// TIA Portal project "IncrocioSemaforicoT" (V19)

(* hardware
DEVICE "S7-1200 station_1"  S7-1200 Station
   slot 0: "Rack_0"  S7-1200 Rack  Rack  V1.0
   slot 1: "PLC_1"  CPU 1212C DC/DC/Rly  6ES7 212-1HE40-0XB0  V4.6
   slot 2: "DQ 16x24VDC_1"  SM 1222 DQ16 x 24VDC  6ES7 222-1BH32-0XB0  V2.0
DEVICE "HMI_1"  KTP700 Basic PN
   slot 0: "HMI_1"  KTP700 Basic PN  6AV2 123-2GB03-0AX0  17.0.0.0
   slot 1: "HMI_RT_1"  KTP700 Basic PN  6AV2 123-2GB03-0AX0  17.0.0.0
   slot 5: "HMI_1.IE_CP_1"  PROFINET Interface  17.0.0.0
      slot 1: "PROFINET Interface_1"  PROFINET Interface
         slot 1: "Port_1"  Port
*)

// ===== PLC "PLC_1"  CPU 1212C DC/DC/Rly =====

VAR_GLOBAL   // PLC tag table "Default tag table"
   "PulsantePedonale1" AT %I0.0 : Bool;
   "PulsantePedonale2" AT %I0.1 : Bool;
   "PulsantePedonale3" AT %I0.2 : Bool;
   "VerdePedonale1" AT %Q0.3 : Bool;
   "GialloPedonale1" AT %Q0.6 : Bool;
   "RossoVeicolare1" AT %Q1.1 : Bool;
   "VerdeVeicolare1" AT %Q1.4 : Bool;
   "GialloVeicolare1" AT %Q1.7 : Bool;
   "RossoPedonale1" AT %Q0.0 : Bool;
   "RossoPedonale2" AT %Q0.1 : Bool;
   "RossoPedonale3" AT %Q0.2 : Bool;
   "VerdePedonale2" AT %Q0.4 : Bool;
   "VerdePedonale3" AT %Q0.5 : Bool;
   "GialloPedonale2" AT %Q0.7 : Bool;
   "GialloPedonale3" AT %Q1.0 : Bool;
   "RossoVeicolare2" AT %Q1.2 : Bool;
   "RossoVeicolare3" AT %Q1.3 : Bool;
   "VerdeVeicolare2" AT %Q1.5 : Bool;
   "VerdeVeicolare3" AT %Q1.6 : Bool;
   "GialloVeicolare2" AT %Q2.0 : Bool;
   "GialloVeicolare3" AT %Q2.1 : Bool;
   "AppoggioGialloVeicolare1" AT %M0.0 : Bool;
   "AppoggioVerdeVeicolare1" AT %M0.1 : Bool;
   "AppoggioQTPRossoVeicolare1" AT %M0.2 : Bool;
   "AppoggioVerdeVeicolare2" AT %M0.3 : Bool;
   "AppoggioGialloVeicolare2" AT %M0.4 : Bool;
   "AppoggioQTPRossoVeicolare2" AT %M0.5 : Bool;
   "AppoggioVerdeVeicolare3" AT %M0.6 : Bool;
   "AppoggioGialloVeicolare3" AT %M0.7 : Bool;
   "AppoggioPulsante1" AT %M1.0 : Bool;
   "AppoggioPulsante2" AT %M1.1 : Bool;
   "AppoggioPulsante3" AT %M1.2 : Bool;
   "AppoggioNVerdePedonale1" AT %M1.3 : Bool;
   "RichiestaPedonale1" AT %M1.4 : Bool;
   "RichiestaPedonale2" AT %M1.5 : Bool;
   "RichiestaPedonale3" AT %M1.6 : Bool;
   "AppoggioPVerdePedonale1" AT %M1.7 : Bool;
   "AppoggioPVerdePedonale2" AT %M2.0 : Bool;
   "AppoggioPVerdePedonale3" AT %M2.1 : Bool;
   "AppoggioQTPRossoVeicolare3" AT %M2.2 : Bool;
   "AppoggioNVerdePedonale2" AT %M2.3 : Bool;
   "AppoggioNVerdePedonale3" AT %M2.4 : Bool;
   "AppoggioQTPRossoVeicolare1Pedonale1" AT %M2.5 : Bool;
   "AppoggioQTPRossoVeicolare1Pedonale3" AT %M2.6 : Bool;
   "AppoggioQTPRossoVeicolare2Pedonale1" AT %M2.7 : Bool;
   "AppoggioQTPRossoVeicolare2Pedonale2" AT %M3.0 : Bool;
   "AppoggioQTPRossoVeicolare3Pedonale2" AT %M3.1 : Bool;
   "AppoggioQTPRossoVeicolare3Pedonale3" AT %M3.2 : Bool;
END_VAR

// folder: System blocks/Program resources

DATA_BLOCK "TPRossoVeicolare1"   // DB1
{ S7_Optimized_Access := 'TRUE' }
AUTHOR : Simatic
FAMILY : IEC
NAME : IEC_TMR
VERSION : 1.0
// stored: InstanceOfName IEC_TIMER
"IEC_TIMER"
BEGIN
END_DATA_BLOCK

DATA_BLOCK "TPVerdeVeicolare1"   // DB2
{ S7_Optimized_Access := 'TRUE' }
AUTHOR : Simatic
FAMILY : IEC
NAME : IEC_TMR
VERSION : 1.0
// stored: InstanceOfName IEC_TIMER
"IEC_TIMER"
BEGIN
END_DATA_BLOCK

DATA_BLOCK "TPGialloVeicolare1"   // DB3
{ S7_Optimized_Access := 'TRUE' }
AUTHOR : Simatic
FAMILY : IEC
NAME : IEC_TMR
VERSION : 1.0
// stored: InstanceOfName IEC_TIMER
"IEC_TIMER"
BEGIN
END_DATA_BLOCK

DATA_BLOCK "TPVerdeVeicolare2"   // DB4
{ S7_Optimized_Access := 'TRUE' }
AUTHOR : Simatic
FAMILY : IEC
NAME : IEC_TMR
VERSION : 1.0
// stored: InstanceOfName IEC_TIMER
"IEC_TIMER"
BEGIN
END_DATA_BLOCK

DATA_BLOCK "TPGialloVeicolare2"   // DB5
{ S7_Optimized_Access := 'TRUE' }
AUTHOR : Simatic
FAMILY : IEC
NAME : IEC_TMR
VERSION : 1.0
// stored: InstanceOfName IEC_TIMER
"IEC_TIMER"
BEGIN
END_DATA_BLOCK

DATA_BLOCK "TPRossoVeicolare2"   // DB6
{ S7_Optimized_Access := 'TRUE' }
AUTHOR : Simatic
FAMILY : IEC
NAME : IEC_TMR
VERSION : 1.0
// stored: InstanceOfName IEC_TIMER
"IEC_TIMER"
BEGIN
END_DATA_BLOCK

DATA_BLOCK "TPVerdeVeicolare3"   // DB7
{ S7_Optimized_Access := 'TRUE' }
AUTHOR : Simatic
FAMILY : IEC
NAME : IEC_TMR
VERSION : 1.0
// stored: InstanceOfName IEC_TIMER
"IEC_TIMER"
BEGIN
END_DATA_BLOCK

DATA_BLOCK "TPGialloVeicolare3"   // DB8
{ S7_Optimized_Access := 'TRUE' }
AUTHOR : Simatic
FAMILY : IEC
NAME : IEC_TMR
VERSION : 1.0
// stored: InstanceOfName IEC_TIMER
"IEC_TIMER"
BEGIN
END_DATA_BLOCK

DATA_BLOCK "TPRossoVeicolare3"   // DB9
{ S7_Optimized_Access := 'TRUE' }
AUTHOR : Simatic
FAMILY : IEC
NAME : IEC_TMR
VERSION : 1.0
// stored: InstanceOfName IEC_TIMER
"IEC_TIMER"
BEGIN
END_DATA_BLOCK

DATA_BLOCK "TPVerdePedonale1"   // DB10
{ S7_Optimized_Access := 'TRUE' }
AUTHOR : Simatic
FAMILY : IEC
NAME : IEC_TMR
VERSION : 1.0
// stored: InstanceOfName IEC_TIMER
"IEC_TIMER"
BEGIN
END_DATA_BLOCK

DATA_BLOCK "TPGialloPedonale1"   // DB11
{ S7_Optimized_Access := 'TRUE' }
AUTHOR : Simatic
FAMILY : IEC
NAME : IEC_TMR
VERSION : 1.0
// stored: InstanceOfName IEC_TIMER
"IEC_TIMER"
BEGIN
END_DATA_BLOCK

DATA_BLOCK "TPVerdePedonale2"   // DB12
{ S7_Optimized_Access := 'TRUE' }
AUTHOR : Simatic
FAMILY : IEC
NAME : IEC_TMR
VERSION : 1.0
// stored: InstanceOfName IEC_TIMER
"IEC_TIMER"
BEGIN
END_DATA_BLOCK

DATA_BLOCK "TPGialloPedonale2"   // DB13
{ S7_Optimized_Access := 'TRUE' }
AUTHOR : Simatic
FAMILY : IEC
NAME : IEC_TMR
VERSION : 1.0
// stored: InstanceOfName IEC_TIMER
"IEC_TIMER"
BEGIN
END_DATA_BLOCK

DATA_BLOCK "TPVerdePedonale3"   // DB14
{ S7_Optimized_Access := 'TRUE' }
AUTHOR : Simatic
FAMILY : IEC
NAME : IEC_TMR
VERSION : 1.0
// stored: InstanceOfName IEC_TIMER
"IEC_TIMER"
BEGIN
END_DATA_BLOCK

DATA_BLOCK "TPGialloPedonale3"   // DB15
{ S7_Optimized_Access := 'TRUE' }
AUTHOR : Simatic
FAMILY : IEC
NAME : IEC_TMR
VERSION : 1.0
// stored: InstanceOfName IEC_TIMER
"IEC_TIMER"
BEGIN
END_DATA_BLOCK

// folder: (top level)

ORGANIZATION_BLOCK "Main"   // OB1, LAD, ProgramCycle
TITLE = "Main Program Sweep (Cycle)"
{ S7_Optimized_Access := 'TRUE' }
VERSION : 0.1
// Incrocio a T con semafori veicolari e pedonali
// 
// A ogni ramo dell'incrocio due semafori veicolari gestiscono attraversamento per immettersi negli altri due rami disponibili: 
// - diventano sincronicamente verdi periodicamente (dopo che lo sono stati quelli su altri rami)
// - siccome le lampade possono essere collegate in parallelo, a livello logico le coppie di semafori (anche pedonali) si possono gestire come singolarità
// 
// I  pedonali, due per ramo, diventano verdi su richiesta, ma solo se i veicolari appartenenti allo stesso ramo sono rossi per ancora almeno 10s. I veicolari sugli altri rami procederanno il loro ciclo indisturbati (le macchine che si devono immettere sul ramo in fase di attraversamento pedonale si fermano in mezzo all'incrocio se trovano occupate le strisce).
// Per fluidificare il traffico e garantire più sicurezza ai pedoni, i pedonali possono diventare verdi solo due volte a ciclo di ramo, ovvero quando scattano i verdi dei veicolari successivi.
// Verde pedonale = 7s
// Giallo pedonale = 3s
// 
// A differenza dei precedenti esercizi semaforici, non è necessario inserire il pulsante di attivazione del ciclo rosso-verde-giallo sui veicolari: il ciclo parte all'avvio della CPU e non si interrompe mai
   VAR_INPUT
      Initial_Call : Bool;   // Initial call of this OB
      Remanence : Bool;   // =True, if remanent data are available
   END_VAR
   VAR_TEMP   // added for the SCL form of the ladder/FBD networks
      _w1 : Bool;
      _w2 : Bool;
      _w3 : Bool;
      _w4 : Bool;
      _w5 : Bool;
   END_VAR
BEGIN

REGION Network 1
   // Veicolare 1
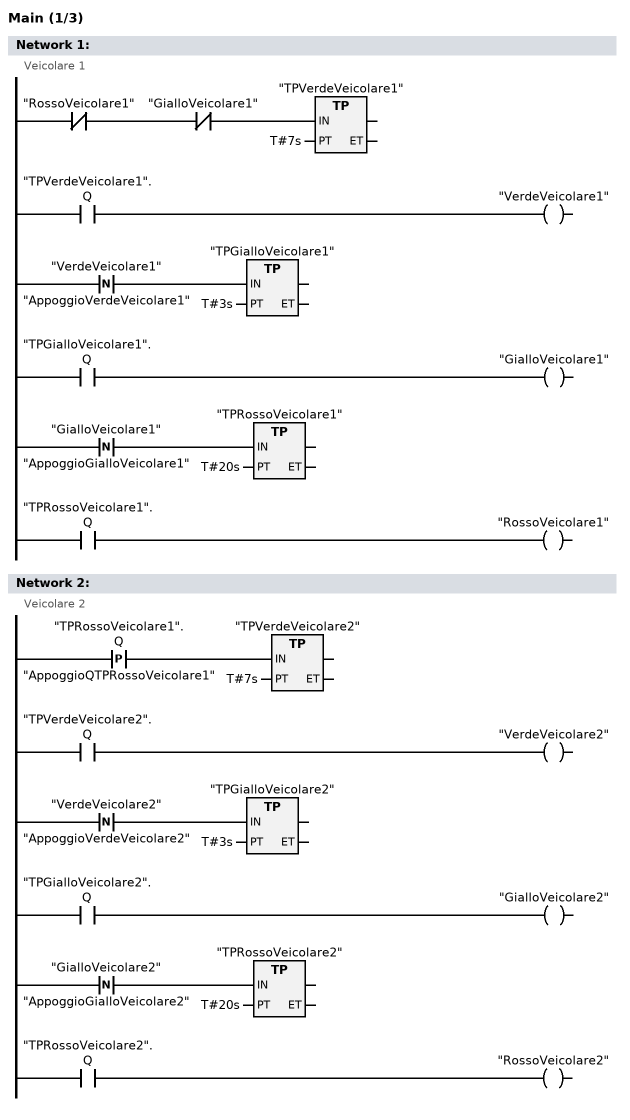
   "TPVerdeVeicolare1".TP(IN := NOT "RossoVeicolare1" AND NOT "GialloVeicolare1", PT := T#7s);
   "VerdeVeicolare1" := "TPVerdeVeicolare1".Q;
   #_w1 := NOT "VerdeVeicolare1" AND "AppoggioVerdeVeicolare1";   // falling edge of "VerdeVeicolare1"
   "AppoggioVerdeVeicolare1" := "VerdeVeicolare1";
   "TPGialloVeicolare1".TP(IN := #_w1, PT := T#3s);
   "GialloVeicolare1" := "TPGialloVeicolare1".Q;
   #_w2 := NOT "GialloVeicolare1" AND "AppoggioGialloVeicolare1";   // falling edge of "GialloVeicolare1"
   "AppoggioGialloVeicolare1" := "GialloVeicolare1";
   "TPRossoVeicolare1".TP(IN := #_w2, PT := T#20s);
   "RossoVeicolare1" := "TPRossoVeicolare1".Q;
END_REGION

REGION Network 2
   // Veicolare 2
   #_w1 := "TPRossoVeicolare1".Q AND NOT "AppoggioQTPRossoVeicolare1";   // rising edge of "TPRossoVeicolare1".Q
   "AppoggioQTPRossoVeicolare1" := "TPRossoVeicolare1".Q;
   "TPVerdeVeicolare2".TP(IN := #_w1, PT := T#7s);
   "VerdeVeicolare2" := "TPVerdeVeicolare2".Q;
   #_w2 := NOT "VerdeVeicolare2" AND "AppoggioVerdeVeicolare2";   // falling edge of "VerdeVeicolare2"
   "AppoggioVerdeVeicolare2" := "VerdeVeicolare2";
   "TPGialloVeicolare2".TP(IN := #_w2, PT := T#3s);
   "GialloVeicolare2" := "TPGialloVeicolare2".Q;
   #_w3 := NOT "GialloVeicolare2" AND "AppoggioGialloVeicolare2";   // falling edge of "GialloVeicolare2"
   "AppoggioGialloVeicolare2" := "GialloVeicolare2";
   "TPRossoVeicolare2".TP(IN := #_w3, PT := T#20s);
   "RossoVeicolare2" := "TPRossoVeicolare2".Q;
END_REGION

REGION Network 3
   // Veicolare 3
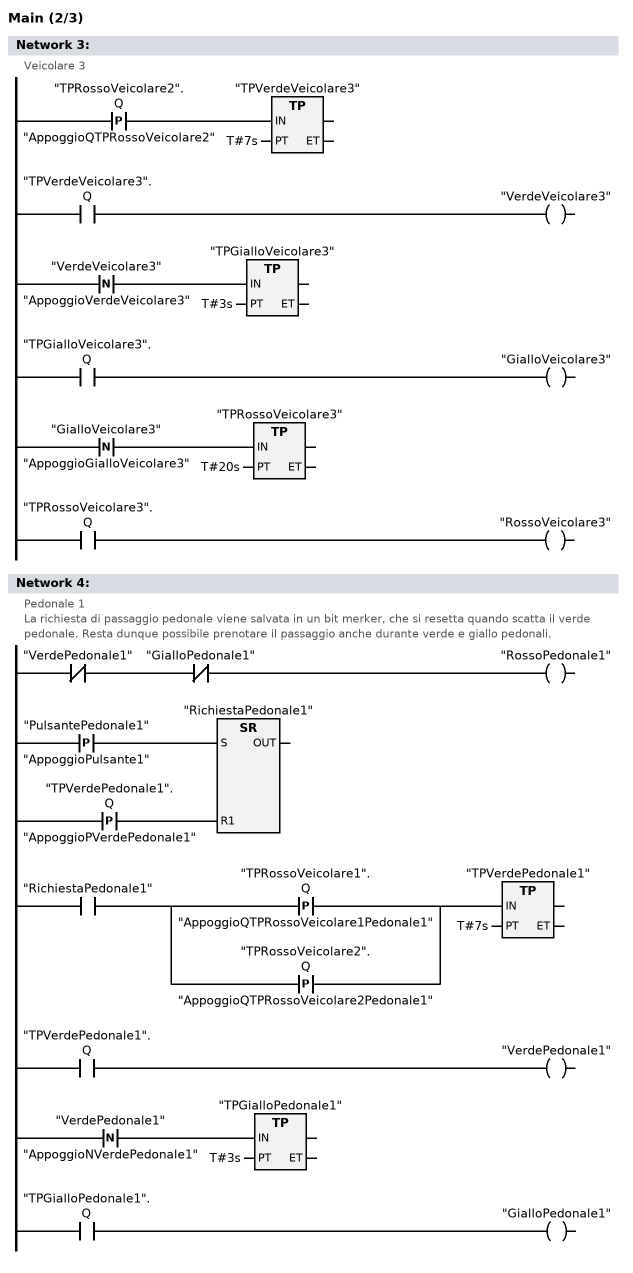
   #_w1 := "TPRossoVeicolare2".Q AND NOT "AppoggioQTPRossoVeicolare2";   // rising edge of "TPRossoVeicolare2".Q
   "AppoggioQTPRossoVeicolare2" := "TPRossoVeicolare2".Q;
   "TPVerdeVeicolare3".TP(IN := #_w1, PT := T#7s);
   "VerdeVeicolare3" := "TPVerdeVeicolare3".Q;
   #_w2 := NOT "VerdeVeicolare3" AND "AppoggioVerdeVeicolare3";   // falling edge of "VerdeVeicolare3"
   "AppoggioVerdeVeicolare3" := "VerdeVeicolare3";
   "TPGialloVeicolare3".TP(IN := #_w2, PT := T#3s);
   "GialloVeicolare3" := "TPGialloVeicolare3".Q;
   #_w3 := NOT "GialloVeicolare3" AND "AppoggioGialloVeicolare3";   // falling edge of "GialloVeicolare3"
   "AppoggioGialloVeicolare3" := "GialloVeicolare3";
   "TPRossoVeicolare3".TP(IN := #_w3, PT := T#20s);
   "RossoVeicolare3" := "TPRossoVeicolare3".Q;
END_REGION

REGION Network 4
   // Pedonale 1
   // 
   // La richiesta di passaggio pedonale viene salvata in un bit merker, che si resetta quando scatta il verde pedonale. Resta dunque possibile prenotare il passaggio anche durante verde e giallo pedonali.
   "RossoPedonale1" := NOT "VerdePedonale1" AND NOT "GialloPedonale1";
   #_w1 := "PulsantePedonale1" AND NOT "AppoggioPulsante1";   // rising edge of "PulsantePedonale1"
   "AppoggioPulsante1" := "PulsantePedonale1";
   #_w2 := "TPVerdePedonale1".Q AND NOT "AppoggioPVerdePedonale1";   // rising edge of "TPVerdePedonale1".Q
   "AppoggioPVerdePedonale1" := "TPVerdePedonale1".Q;
   IF #_w1 THEN
       "RichiestaPedonale1" := TRUE;   // SR flip-flop
   END_IF;
   IF #_w2 THEN "RichiestaPedonale1" := FALSE; END_IF;
   #_w3 := "RichiestaPedonale1" AND "TPRossoVeicolare1".Q AND NOT "AppoggioQTPRossoVeicolare1Pedonale1";   // rising edge of "TPRossoVeicolare1".Q
   "AppoggioQTPRossoVeicolare1Pedonale1" := "TPRossoVeicolare1".Q;
   #_w4 := "RichiestaPedonale1" AND "TPRossoVeicolare2".Q AND NOT "AppoggioQTPRossoVeicolare2Pedonale1";   // rising edge of "TPRossoVeicolare2".Q
   "AppoggioQTPRossoVeicolare2Pedonale1" := "TPRossoVeicolare2".Q;
   "TPVerdePedonale1".TP(IN := #_w3 OR #_w4, PT := T#7s);
   "VerdePedonale1" := "TPVerdePedonale1".Q;
   #_w5 := NOT "VerdePedonale1" AND "AppoggioNVerdePedonale1";   // falling edge of "VerdePedonale1"
   "AppoggioNVerdePedonale1" := "VerdePedonale1";
   "TPGialloPedonale1".TP(IN := #_w5, PT := T#3s);
   "GialloPedonale1" := "TPGialloPedonale1".Q;
END_REGION

REGION Network 5
   // Pedonale 2
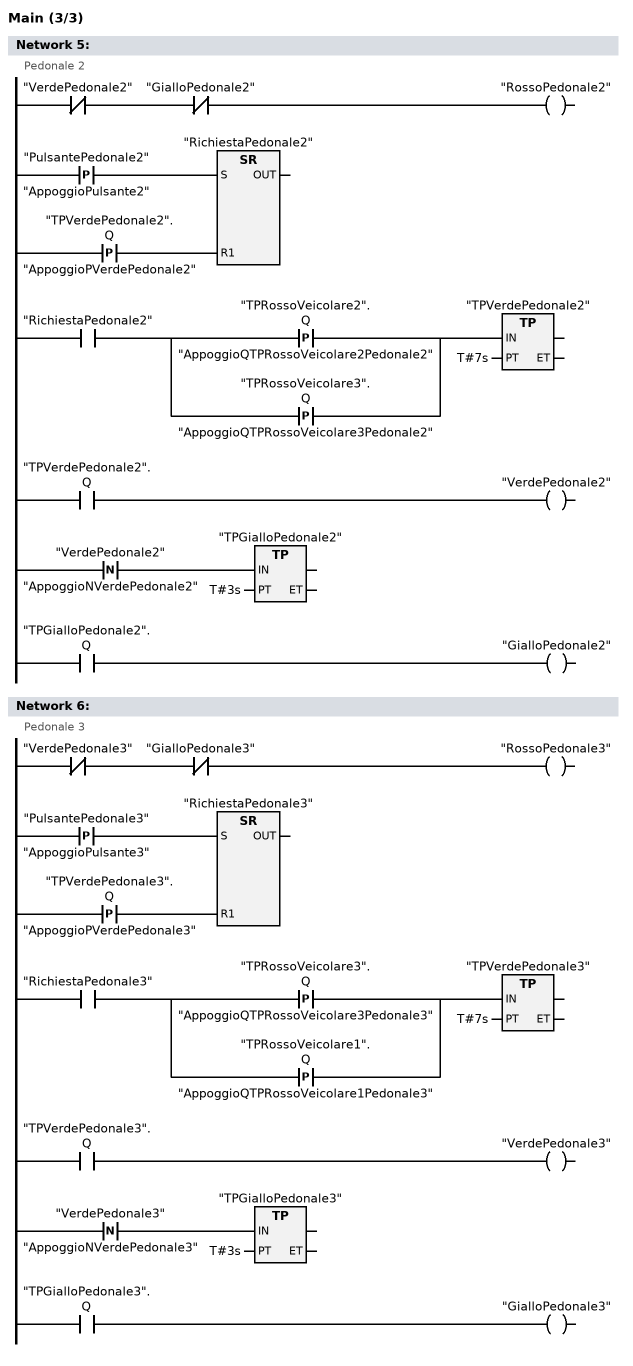
   "RossoPedonale2" := NOT "VerdePedonale2" AND NOT "GialloPedonale2";
   #_w1 := "PulsantePedonale2" AND NOT "AppoggioPulsante2";   // rising edge of "PulsantePedonale2"
   "AppoggioPulsante2" := "PulsantePedonale2";
   #_w2 := "TPVerdePedonale2".Q AND NOT "AppoggioPVerdePedonale2";   // rising edge of "TPVerdePedonale2".Q
   "AppoggioPVerdePedonale2" := "TPVerdePedonale2".Q;
   IF #_w1 THEN
       "RichiestaPedonale2" := TRUE;   // SR flip-flop
   END_IF;
   IF #_w2 THEN "RichiestaPedonale2" := FALSE; END_IF;
   #_w3 := "RichiestaPedonale2" AND "TPRossoVeicolare2".Q AND NOT "AppoggioQTPRossoVeicolare2Pedonale2";   // rising edge of "TPRossoVeicolare2".Q
   "AppoggioQTPRossoVeicolare2Pedonale2" := "TPRossoVeicolare2".Q;
   #_w4 := "RichiestaPedonale2" AND "TPRossoVeicolare3".Q AND NOT "AppoggioQTPRossoVeicolare3Pedonale2";   // rising edge of "TPRossoVeicolare3".Q
   "AppoggioQTPRossoVeicolare3Pedonale2" := "TPRossoVeicolare3".Q;
   "TPVerdePedonale2".TP(IN := #_w3 OR #_w4, PT := T#7s);
   "VerdePedonale2" := "TPVerdePedonale2".Q;
   #_w5 := NOT "VerdePedonale2" AND "AppoggioNVerdePedonale2";   // falling edge of "VerdePedonale2"
   "AppoggioNVerdePedonale2" := "VerdePedonale2";
   "TPGialloPedonale2".TP(IN := #_w5, PT := T#3s);
   "GialloPedonale2" := "TPGialloPedonale2".Q;
END_REGION

REGION Network 6
   // Pedonale 3
   "RossoPedonale3" := NOT "VerdePedonale3" AND NOT "GialloPedonale3";
   #_w1 := "PulsantePedonale3" AND NOT "AppoggioPulsante3";   // rising edge of "PulsantePedonale3"
   "AppoggioPulsante3" := "PulsantePedonale3";
   #_w2 := "TPVerdePedonale3".Q AND NOT "AppoggioPVerdePedonale3";   // rising edge of "TPVerdePedonale3".Q
   "AppoggioPVerdePedonale3" := "TPVerdePedonale3".Q;
   IF #_w1 THEN
       "RichiestaPedonale3" := TRUE;   // SR flip-flop
   END_IF;
   IF #_w2 THEN "RichiestaPedonale3" := FALSE; END_IF;
   #_w3 := "RichiestaPedonale3" AND "TPRossoVeicolare3".Q AND NOT "AppoggioQTPRossoVeicolare3Pedonale3";   // rising edge of "TPRossoVeicolare3".Q
   "AppoggioQTPRossoVeicolare3Pedonale3" := "TPRossoVeicolare3".Q;
   #_w4 := "RichiestaPedonale3" AND "TPRossoVeicolare1".Q AND NOT "AppoggioQTPRossoVeicolare1Pedonale3";   // rising edge of "TPRossoVeicolare1".Q
   "AppoggioQTPRossoVeicolare1Pedonale3" := "TPRossoVeicolare1".Q;
   "TPVerdePedonale3".TP(IN := #_w3 OR #_w4, PT := T#7s);
   "VerdePedonale3" := "TPVerdePedonale3".Q;
   #_w5 := NOT "VerdePedonale3" AND "AppoggioNVerdePedonale3";   // falling edge of "VerdePedonale3"
   "AppoggioNVerdePedonale3" := "VerdePedonale3";
   "TPGialloPedonale3".TP(IN := #_w5, PT := T#3s);
   "GialloPedonale3" := "TPGialloPedonale3".Q;
END_REGION
END_ORGANIZATION_BLOCK

(* ===== HMI "HMI_RT_1" =====
system functions are stored by id; their names below are inferred from use
connection "HMI_Connection_1": ETHERNET, SMART_S7_1200_OMS

HMI tags "Default tag table"
   "Tag_ScreenNumber" : UInt, internal
   "PulsantePedonale3" : Bool = PLC PulsantePedonale3 AT %I0.2, 100 ms
   "PulsantePedonale1" : Bool = PLC PulsantePedonale1 AT %I0.0, 100 ms
   "PulsantePedonale2" : Bool = PLC PulsantePedonale2 AT %I0.1, 100 ms
   "VerdePedonale3" : Bool = PLC VerdePedonale3 AT %Q0.5, 100 ms
   "RossoPedonale3" : Bool = PLC RossoPedonale3 AT %Q0.2, 100 ms
   "GialloPedonale3" : Bool = PLC GialloPedonale3 AT %Q1.0, 100 ms
   "RossoPedonale1" : Bool = PLC RossoPedonale1 AT %Q0.0, 100 ms
   "GialloPedonale1" : Bool = PLC GialloPedonale1 AT %Q0.6, 100 ms
   "VerdePedonale1" : Bool = PLC VerdePedonale1 AT %Q0.3, 100 ms
   "RossoPedonale2" : Bool = PLC RossoPedonale2 AT %Q0.1, 100 ms
   "GialloPedonale2" : Bool = PLC GialloPedonale2 AT %Q0.7, 100 ms
   "VerdePedonale2" : Bool = PLC VerdePedonale2 AT %Q0.4, 100 ms
   "RossoVeicolare1" : Bool = PLC RossoVeicolare1 AT %Q1.1, 100 ms
   "GialloVeicolare1" : Bool = PLC GialloVeicolare1 AT %Q1.7, 100 ms
   "VerdeVeicolare1" : Bool = PLC VerdeVeicolare1 AT %Q1.4, 100 ms
   "RossoVeicolare2" : Bool = PLC RossoVeicolare2 AT %Q1.2, 100 ms
   "GialloVeicolare2" : Bool = PLC GialloVeicolare2 AT %Q2.0, 100 ms
   "VerdeVeicolare2" : Bool = PLC VerdeVeicolare2 AT %Q1.5, 100 ms
   "RossoVeicolare3" : Bool = PLC RossoVeicolare3 AT %Q1.3, 100 ms
   "GialloVeicolare3" : Bool = PLC GialloVeicolare3 AT %Q2.1, 100 ms
   "VerdeVeicolare3" : Bool = PLC VerdeVeicolare3 AT %Q1.6, 100 ms
   "RichiestaPedonale2" : Bool = PLC RichiestaPedonale2 AT %M1.5, 1 s
   "RichiestaPedonale1" : Bool = PLC RichiestaPedonale1 AT %M1.4, 1 s
   "RichiestaPedonale3" : Bool = PLC RichiestaPedonale3 AT %M1.6, 1 s

Template "Template_1" 800x480
   Button "Exit" at 714,429 size 71x50; TextOff 'Exit'; PictureOff "ExitRuntime_KTP700_Basic_PN_TR"; PictureOn "ExitRuntime_KTP700_Basic_PN_TR"
      on Release: StopRuntime(0)
   Button "Language" at 614,429 size 71x50; TextOff 'Language'; PictureOff "ToggleLanguage_KTP700_Basic_PN_TR"; PictureOn "ToggleLanguage_KTP700_Basic_PN_TR"
      on Release: function_fb9197e8(-1)
   Button "Log on" at 514,429 size 71x50; TextOff 'Log on'; PictureOff "Login_KTP700_Basic_PN_TR"; PictureOn "Login_KTP700_Basic_PN_TR"
      on Release: function_a2a04561()
   Button "Template_Button" at 414,429 size 71x50; TextOff 'Text'
   Button "Template_Button_1" at 314,429 size 71x50; TextOff 'Text'
   Button "Template_Button_2" at 214,429 size 71x50; TextOff 'Text'
   Button "Alarms" at 114,429 size 71x50; TextOff 'Alarms'; PictureOff "AlarmDisplay_KTP700_Basic_PN_TR"; PictureOn "AlarmDisplay_KTP700_Basic_PN_TR"
      on Release: function_ef3f5d25("Alarm window_Unacknowledged", -1)
   Button "Start screen" at 14,429 size 71x50; TextOff 'Start screen'; PictureOff "NavigateHome_KTP700_Basic_PN_TR"; PictureOn "NavigateHome_KTP700_Basic_PN_TR"
      on Release: ActivateScreen("Incrocio", 0)
   SymbolicIOField "Symbolic_IO_Field_Screen" at 53,9 size 640x33; TextOff '0'; TextOn '1'; TextList "TextList_ScreenNames"
      ProcessValue <- "Tag_ScreenNumber"
      on Change: ActivateScreenByNumber("Tag_ScreenNumber", 0)
   DateTimeField "HmiScreenItemData" at 695,25 size 105x25
   DateTimeField "HmiScreenItemData_1" at 695,0 size 105x25
   GraphicView "Logo" at 0,0 size 51x51; Picture "Logo of HMI_1"

screen "Incrocio" 800x480, template "Template_1"
   on GenerateScreen: SetTag("Tag_ScreenNumber", 1)
   Button "HmiScreenItemData" at 173,50 size 159x47; TextOff 'Ramo 1'; PictureOff "Navigates to Ramo 1 for KTP700 Basic+ PN 17.0.0.0"; PictureOn "Navigates to Ramo 1 for KTP700 Basic+ PN 17.0.0.0"
      on Release: ActivateScreen("Ramo 1", 0)
   Button "HmiScreenItemData_1" at 333,50 size 159x47; TextOff 'Ramo 2'; PictureOff "Navigates to Ramo 2 for KTP700 Basic+ PN 17.0.0.0"; PictureOn "Navigates to Ramo 2 for KTP700 Basic+ PN 17.0.0.0"
      on Release: ActivateScreen("Ramo 2", 0)
   Button "HmiScreenItemData_2" at 493,50 size 159x47; TextOff 'Ramo 3'; PictureOff "Navigates to Ramo 3 for KTP700 Basic+ PN 17.0.0.0"; PictureOn "Navigates to Ramo 3 for KTP700 Basic+ PN 17.0.0.0"
      on Release: ActivateScreen("Ramo 3", 0)
   Button "HmiScreenItemData_4" at 285,431 size 159x47; TextOff 'System screens'; PictureOff "Navigates to System screens for KTP700 Basic+ PN 17.0.0.0"; PictureOn "Navigates to System screens for KTP700 Basic+ PN 17.0.0.0"
      on Release: ActivateScreen("System screens", 0)
   GraphicView "Graphic view_1" at 16,104 size 771x315; Picture "BgHMI"
   Group "Group_5" at 49,295 size 45x104
   GraphicView "Graphic view_2" at 671,141 size 75x147; Picture "PedonaliBgHMI"
   GraphicView "Graphic view_4" at 226,350 size 236x60; Picture "PedonaliOrizBgHMI"
   Button "Button_1" at 658,107 size 99x32; TextOff 'Richiesta 2'
      on Press: SetBit("RichiestaPedonale2")
   Button "Button_2" at 21,107 size 99x32; TextOff 'Richiesta 3'
      on Press: SetBit("RichiestaPedonale3")
   Button "Button_4" at 122,380 size 99x32; TextOff 'Richiesta 1'
      on Press: SetBit("RichiestaPedonale1")
   Group "Group_1" at 201,191 size 45x104
   Group "Group_2" at 466,309 size 45x104
   Group "Group_3" at 685,295 size 45x104
   Group "Group_4" at 444,110 size 45x104
   Group "Group_6" at 383,237 size 45x104
   Button "FB_Empty_Round" at 514,309 size 50x50; TextOff 'Text'; PictureOff "FB_Empty_Round_Released_256c"; PictureOn "FB_Empty_Round_Pressed_256c"
      on Press: SetBit("RichiestaPedonale1")
   Button "FB_Empty_Round_1" at 633,295 size 50x50; TextOff 'Text'; PictureOff "FB_Empty_Round_Released_256c"; PictureOn "FB_Empty_Round_Pressed_256c"
      on Press: SetBit("RichiestaPedonale2")
   Button "FB_Empty_Round_2" at 99,295 size 50x50; TextOff 'Text'; PictureOff "FB_Empty_Round_Released_256c"; PictureOn "FB_Empty_Round_Pressed_256c"
      on Press: SetBit("RichiestaPedonale3")
   GraphicView "Graphic view_3" at 35,141 size 75x147; Picture "PedonaliBgHMI"
   Circle "Circle_16" at 57,298 size 29x29
      Appearance <- "RossoPedonale3"
   Circle "Circle_17" at 57,332 size 29x29
      Appearance <- "GialloPedonale3"
   Circle "Circle_18" at 57,366 size 29x29
      Appearance <- "VerdePedonale3"
   Circle "Circle_1" at 209,194 size 29x29
      Appearance <- "RossoVeicolare3"
   Circle "Circle_2" at 209,228 size 29x29
      Appearance <- "GialloVeicolare3"
   Circle "Circle_3" at 209,262 size 29x29
      Appearance <- "VerdeVeicolare3"
   Circle "Circle_4" at 474,312 size 29x29
      Appearance <- "RossoPedonale1"
   Circle "Circle_5" at 474,346 size 29x29
      Appearance <- "GialloPedonale1"
   Circle "Circle_6" at 474,380 size 29x29
      Appearance <- "VerdePedonale1"
   Circle "Circle_7" at 693,298 size 29x29
      Appearance <- "RossoPedonale2"
   Circle "Circle_8" at 693,332 size 29x29
      Appearance <- "GialloPedonale2"
   Circle "Circle_9" at 693,366 size 29x29
      Appearance <- "VerdePedonale2"
   Circle "Circle_10" at 452,113 size 29x29
      Appearance <- "RossoVeicolare2"
   Circle "Circle_11" at 452,147 size 29x29
      Appearance <- "GialloVeicolare2"
   Circle "Circle_12" at 452,181 size 29x29
      Appearance <- "VerdeVeicolare2"
   Circle "Circle_13" at 391,240 size 29x29
      Appearance <- "RossoVeicolare1"
   Circle "Circle_14" at 391,274 size 29x29
      Appearance <- "GialloVeicolare1"
   Circle "Circle_15" at 391,308 size 29x29
      Appearance <- "VerdeVeicolare1"

screen "Ramo 1" 800x480, template "Template_1"
   on GenerateScreen: SetTag("Tag_ScreenNumber", 2)
   TextField "HmiScreenItemData" at 80,225 size 640x25; Text 'Ramo 1'
   Button "Back" at 1,52 size 159x47; TextOff 'Back'
      on Release: ActivateScreen("Incrocio", 0)
   Button "HmiScreenItemData_1" at 36,146 size 159x47; TextOff 'Veicolare 1'; PictureOff "Navigates to Veicolare 1 for KTP700 Basic+ PN 17.0.0.0"; PictureOn "Navigates to Veicolare 1 for KTP700 Basic+ PN 17.0.0.0"
      on Release: ActivateScreen("Veicolare 1", 0)
   Button "HmiScreenItemData_2" at 36,205 size 159x47; TextOff 'Pedonale 1'; PictureOff "Navigates to Pedonale 1 for KTP700 Basic+ PN 17.0.0.0"; PictureOn "Navigates to Pedonale 1 for KTP700 Basic+ PN 17.0.0.0"
      on Release: ActivateScreen("Pedonale 1", 0)

screen "Veicolare 1" 800x480, template "Template_1"
   on GenerateScreen: SetTag("Tag_ScreenNumber", 3)
   TextField "HmiScreenItemData" at 80,225 size 640x25; Text 'Veicolare 1'
   Button "Back" at 1,52 size 159x47; TextOff 'Back'
      on Release: ActivateScreen("Ramo 1", 0)

screen "Pedonale 1" 800x480, template "Template_1"
   on GenerateScreen: SetTag("Tag_ScreenNumber", 4)
   TextField "HmiScreenItemData" at 80,225 size 640x25; Text 'Pedonale 1'
   Button "Back" at 268,431 size 159x47; TextOff 'Back'
      on Release: ActivateScreen("Ramo 1", 0)
   HTMLBrowser "HTML browser_1" at 18,50 size 764x372

screen "Ramo 2" 800x480, template "Template_1"
   on GenerateScreen: SetTag("Tag_ScreenNumber", 5)
   TextField "HmiScreenItemData" at 80,225 size 640x25; Text 'Ramo 2'
   Button "Back" at 1,52 size 159x47; TextOff 'Back'
      on Release: ActivateScreen("Incrocio", 0)
   Button "HmiScreenItemData_1" at 36,146 size 159x47; TextOff 'Veicolare 2'; PictureOff "Navigates to Veicolare 2 for KTP700 Basic+ PN 17.0.0.0"; PictureOn "Navigates to Veicolare 2 for KTP700 Basic+ PN 17.0.0.0"
      on Release: ActivateScreen("Veicolare 2", 0)
   Button "HmiScreenItemData_2" at 36,205 size 159x47; TextOff 'Pedonale 2'; PictureOff "Navigates to Pedonale 2 for KTP700 Basic+ PN 17.0.0.0"; PictureOn "Navigates to Pedonale 2 for KTP700 Basic+ PN 17.0.0.0"
      on Release: ActivateScreen("Pedonale 2", 0)

screen "Veicolare 2" 800x480, template "Template_1"
   on GenerateScreen: SetTag("Tag_ScreenNumber", 6)
   TextField "HmiScreenItemData" at 80,225 size 640x25; Text 'Veicolare 2'
   Button "Back" at 1,52 size 159x47; TextOff 'Back'
      on Release: ActivateScreen("Ramo 2", 0)

screen "Pedonale 2" 800x480, template "Template_1"
   on GenerateScreen: SetTag("Tag_ScreenNumber", 7)
   TextField "HmiScreenItemData" at 80,225 size 640x25; Text 'Pedonale 2'
   Button "Back" at 1,52 size 159x47; TextOff 'Back'
      on Release: ActivateScreen("Ramo 2", 0)

screen "Ramo 3" 800x480, template "Template_1"
   on GenerateScreen: SetTag("Tag_ScreenNumber", 8)
   TextField "HmiScreenItemData" at 80,225 size 640x25; Text 'Ramo 3'
   Button "Back" at 1,52 size 159x47; TextOff 'Back'
      on Release: ActivateScreen("Incrocio", 0)
   Button "HmiScreenItemData_1" at 36,146 size 159x47; TextOff 'Veicolare 3'; PictureOff "Navigates to Veicolare 3 for KTP700 Basic+ PN 17.0.0.0"; PictureOn "Navigates to Veicolare 3 for KTP700 Basic+ PN 17.0.0.0"
      on Release: ActivateScreen("Veicolare 3", 0)
   Button "HmiScreenItemData_2" at 36,205 size 159x47; TextOff 'Pedonale 3'; PictureOff "Navigates to Pedonale 3 for KTP700 Basic+ PN 17.0.0.0"; PictureOn "Navigates to Pedonale 3 for KTP700 Basic+ PN 17.0.0.0"
      on Release: ActivateScreen("Pedonale 3", 0)

screen "Veicolare 3" 800x480, template "Template_1"
   on GenerateScreen: SetTag("Tag_ScreenNumber", 9)
   TextField "HmiScreenItemData" at 80,225 size 640x25; Text 'Veicolare 3'
   Button "Back" at 1,52 size 159x47; TextOff 'Back'
      on Release: ActivateScreen("Ramo 3", 0)

screen "Pedonale 3" 800x480, template "Template_1"
   on GenerateScreen: SetTag("Tag_ScreenNumber", 10)
   TextField "HmiScreenItemData" at 80,225 size 640x25; Text 'Pedonale 3'
   Button "Back" at 1,52 size 159x47; TextOff 'Back'
      on Release: ActivateScreen("Ramo 3", 0)

screen "System screens" 800x480, template "Template_1"
   on GenerateScreen: SetTag("Tag_ScreenNumber", 11)
   Button "Back" at 1,52 size 159x47; TextOff 'Back'
      on Release: ActivateScreen("Incrocio", 0)
   Button "HmiScreenItemData" at 36,146 size 159x47; TextOff 'Different jobs'; PictureOff "Navigates to Different jobs for KTP700 Basic+ PN 17.0.0.0"; PictureOn "Navigates to Different jobs for KTP700 Basic+ PN 17.0.0.0"
      on Release: ActivateScreen("Different jobs", 0)

screen "Different jobs" 800x480, template "Template_1"
   on GenerateScreen: SetTag("Tag_ScreenNumber", 12)
   Button "Online" at 36,146 size 159x47; TextOff 'Online'
      on Release: function_bb44b551(0)
   Button "Offline" at 36,205 size 159x47; TextOff 'Offline'
      on Release: function_bb44b551(1)
   Button "Transfer" at 36,264 size 159x47; TextOff 'Transfer'
      on Release: function_bb44b551(2)
   Button "Toggle language" at 36,323 size 159x47; TextOff 'Toggle language'
      on Release: function_fb9197e8(-1)
   Button "Stop Runtime" at 207,146 size 159x47; TextOff 'Stop Runtime'
      on Release: StopRuntime(0)
   Button "Back" at 1,52 size 159x47; TextOff 'Back'
      on Release: ActivateScreen("System screens", 0)
*)